(* IEC 61131-3 sources: codesys-to-s7/tests/fixtures/s7-to-codesys/src/DUTs/Converted, 7 files *)

(* ---- ST_DB_Hmi_pump.dut.st ---- *)
// Назначение: структура поля «pump» блока «DB_Hmi» (анонимный Struct в SCL)
// Автор:      s7conv 0.1.0 (сгенерировано)
// Версия:     не указана
// Документ:   docs/MAPPING.md, раздел «Типы»
// Источник:   samples/scl/DB_Plant.scl, DATA_BLOCK "DB_Hmi"
TYPE ST_DB_Hmi_pump :
STRUCT
    // Команды насосам P101...P103
    startReq : BOOL;
    stopReq : BOOL;
    resetReq : BOOL;
END_STRUCT
END_TYPE

(* ---- ST_DB_Plant_shiftData.dut.st ---- *)
// Назначение: структура поля «shiftData» блока «DB_Plant» (анонимный Struct в SCL)
// Автор:      s7conv 0.1.0 (сгенерировано)
// Версия:     не указана
// Документ:   docs/MAPPING.md, раздел «Типы»
// Источник:   samples/scl/DB_Plant.scl, DATA_BLOCK "DB_Plant"
TYPE ST_DB_Plant_shiftData :
STRUCT
    // Данные смены
    startedAt : DT;  // Начало смены
    volume : LREAL;  // Объём за смену, м3
    pumpStarts : DINT;  // Пуски насосов за смену
END_STRUCT
END_TYPE

(* ---- ST_FB_EventLogger_buffer.dut.st ---- *)
// Назначение: структура поля «buffer» блока «FB_EventLogger» (анонимный Struct в SCL)
// Автор:      s7conv 0.1.0 (сгенерировано)
// Версия:     не указана
// Документ:   docs/MAPPING.md, раздел «Типы»
// Источник:   samples/scl/FB_EventLogger.scl, FUNCTION_BLOCK "FB_EventLogger"
TYPE ST_FB_EventLogger_buffer :
STRUCT
    // Кольцевой буфер
    stamp : DT;
    code : INT;
    aux : INT;
    text : STRING(20);
END_STRUCT
END_TYPE

(* ---- ST_UDT_AnalogCfg_limits.dut.st ---- *)
// Назначение: структура поля «limits» блока «UDT_AnalogCfg» (анонимный Struct в SCL)
// Автор:      s7conv 0.1.0 (сгенерировано)
// Версия:     не указана
// Документ:   docs/MAPPING.md, раздел «Типы»
// Источник:   samples/scl/UDT_PlantTypes.scl, TYPE "UDT_AnalogCfg"
TYPE ST_UDT_AnalogCfg_limits :
STRUCT
    // Уставки сигнализации, инж. ед.
    hh : REAL := 14.0;  // Аварийно высокое
    h : REAL := 12.0;  // Предупредительно высокое
    l : REAL := 2.0;  // Предупредительно низкое
    ll : REAL := 1.0;  // Аварийно низкое
END_STRUCT
END_TYPE

(* ---- UDT_AnalogCfg.dut.st ---- *)
// Назначение: Тип (UDT) «UDT_AnalogCfg», сконвертирован из SCL
// Автор:      не указан (исходный блок S7); перевод в ST — s7conv 0.1.0
// Версия:     0.1 (исходный блок S7)
// Документ:   docs/CONVERSION_REPORT.md, docs/MAPPING.md
// Источник:   samples/scl/UDT_PlantTypes.scl, строки 23–38, TYPE "UDT_AnalogCfg"
// Сгенерировано s7conv: пометки MIGRATION-CHECK и MIGRATION-TODO требуют ручного разбора.
// ---- комментарий в начале исходного файла SCL ----
// =============================================================================
// s7-to-codesys — корпус SCL. Написан с нуля для проекта, это не выгрузка
// реального объекта. Вымышленный объект: ВОС «Северная» — насосная станция
// II подъёма, скорые фильтры, дозирование реагента.
//
// Файл:   UDT_PlantTypes.scl
// Блоки:  TYPE "UDT_AnalogCfg", TYPE "UDT_DeviceStatus", TYPE "UDT_DosingRecipe"
// -----------------------------------------------------------------------------
// Назначение
//   Пользовательские типы данных (PLC data types) станции. Логики нет.
//   UDT_AnalogCfg    — параметры аналогового канала: шкала, уставки (вложенная
//                      структура limits), гистерезис, единица измерения.
//   UDT_DeviceStatus — состояние устройства для HMI: работа, авария, режим,
//                      код аварии, число пусков. Его заполняет FB_Motor.
//   UDT_DosingRecipe — рецепт дозирования: имя (String[20]), реагент, дозы по
//                      ступеням (Array[1..4] of Real), время контакта (Time),
//                      отметка изменения (Date_And_Time), признак утверждения.
// Что проверяет при конвертации
//   TYPE/STRUCT/END_STRUCT; вложенная анонимная Struct; массив в структуре с
//   инициализатором [..] и множителем повторения; значения по умолчанию;
//   String[n] -> STRING(n); Date_And_Time -> DT; Time -> TIME.
// =============================================================================
TYPE UDT_AnalogCfg :
STRUCT
    rangeLow : REAL := 0.0;  // Значение при raw = 0, инж. ед.
    rangeHigh : REAL := 16.0;  // Значение при raw = 27648, инж. ед.
    limits : ST_UDT_AnalogCfg_limits;
    hysteresis : REAL := 0.5;  // Гистерезис уставок, инж. ед.
    unitText : STRING(8) := 'bar';  // Единица измерения для HMI
END_STRUCT
END_TYPE

(* ---- UDT_DeviceStatus.dut.st ---- *)
// Назначение: Тип (UDT) «UDT_DeviceStatus», сконвертирован из SCL
// Автор:      не указан (исходный блок S7); перевод в ST — s7conv 0.1.0
// Версия:     0.1 (исходный блок S7)
// Документ:   docs/CONVERSION_REPORT.md, docs/MAPPING.md
// Источник:   samples/scl/UDT_PlantTypes.scl, строки 40–50, TYPE "UDT_DeviceStatus"
// Сгенерировано s7conv: пометки MIGRATION-CHECK и MIGRATION-TODO требуют ручного разбора.
TYPE UDT_DeviceStatus :
STRUCT
    running : BOOL;  // Работает (команда и обратная связь)
    fault : BOOL;  // Авария (защёлка)
    autoMode : BOOL;  // Режим авто
    faultCode : INT;  // 0 — нет, 1 — нет ОС после пуска, 2 — пропала ОС, 3 — тепловая защита, 4 — ОС без команды
    startCount : DINT;  // Число пусков
END_STRUCT
END_TYPE

(* ---- UDT_DosingRecipe.dut.st ---- *)
// Назначение: Тип (UDT) «UDT_DosingRecipe», сконвертирован из SCL
// Автор:      не указан (исходный блок S7); перевод в ST — s7conv 0.1.0
// Версия:     0.2 (исходный блок S7)
// Документ:   docs/CONVERSION_REPORT.md, docs/MAPPING.md
// Источник:   samples/scl/UDT_PlantTypes.scl, строки 52–64, TYPE "UDT_DosingRecipe"
// Сгенерировано s7conv: пометки MIGRATION-CHECK и MIGRATION-TODO требуют ручного разбора.
TYPE UDT_DosingRecipe :
STRUCT
    name : STRING(20) := 'DEFAULT';  // Имя рецепта
    reagent : INT := 1;  // 1 — коагулянт, 2 — флокулянт, 3 — гипохлорит
    doseStep : ARRAY[1..4] OF REAL := [0.5, 1.0, 1.5, 2.0];  // Доза по ступеням расхода, мг/л
    stepFlow : ARRAY[1..4] OF REAL := [4(0.0)];  // Границы ступеней расхода, м3/ч (задаются с HMI)
    contactTime : TIME := T#15M;  // Время контакта
    changedAt : DT := DT#2024-01-01-00:00:00;  // Когда изменён
    approved : BOOL;  // Утверждён технологом
END_STRUCT
END_TYPE
